Fanuc KAREL source: ko00100.KL

-- PROVISIONAL review KL for V770-1; original PC SHA256 3866f11bc9163d489fc93fd3cae345f7cbb995553b0998fa0b7dc8baba6ec820
-- Incomplete behavior may be omitted. Consult companion uncertainty JSON. Do not deploy.
PROGRAM KO00100
%NOLOCKGROUP
VAR
  A : INTEGER
  B : REAL
  OUT : REAL
BEGIN
  -- UNRESOLVED_PC offsets 5-12; opcodes 9D,23
  -- UNRESOLVED_PC offsets 17-29; opcodes 2E,64,23
  -- UNRESOLVED_PC offsets 34-57; opcodes 27,27,21,64,22,76,23
  -- UNRESOLVED_PC offsets 62-66; opcodes 7F
END KO00100
